// TIA Portal V21 export
// export: Created 2026-11-11T00:47:14.8809745Z, ExportSetting WithDefaults, DisplayName Totally Integrated Automation Portal, DisplayVersion V21 Update 3, DisplayName STEP 7 Professional, DisplayVersion V21 Update 3, DisplayName STEP 7 Safety, DisplayVersion V21, DisplayName Tech WebApplication, DisplayVersion V21, DisplayName WinCC Basic/Comfort/Advanced, DisplayVersion V21 Update 3, DisplayName WinCC Unified, DisplayVersion V21 Update 3
FUNCTION_BLOCK "FB_Fbd_ex037"   // FB360, FBD
{ S7_Optimized_Access := 'TRUE' }
VERSION : 0.1
// stored: AutoNumber true, IsIECCheckEnabled false, IsRetainMemResEnabled false, MemoryReserve 100, SetENOAutomatically false, UDAEnableTagReadback false
   VAR_INPUT
      v_size : DInt;
   END_VAR
   VAR_OUTPUT
      v_out : WString;
   END_VAR
   VAR_IN_OUT
      v_variable : Variant;
   END_VAR
BEGIN

REGION Network 1: Querying GetSymbolPath - actual parameter at beginning of a call path
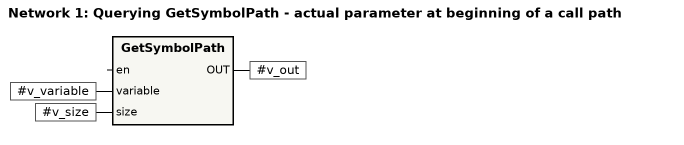
   GetSymbolPath(variable := #v_variable, size := #v_size, OUT => #v_out);
END_REGION
END_FUNCTION_BLOCK
